{attribute 'no_assign'}
FUNCTION_BLOCK FB_DO_WTURBINE_LD0_LLN0_NamPlt EXTENDS FB_AcsiCommonDataClass
VAR_INPUT
	vendor: FB_AcsiDATypeVisString255 := (Fc:=ACSI_FC_DC, bLinkResult:=THIS^.AddDataToContainer(ipData:=vendor));
	swRev: FB_AcsiDATypeVisString255 := (Fc:=ACSI_FC_DC, bLinkResult:=THIS^.AddDataToContainer(ipData:=swRev));
	ldNs: FB_AcsiDATypeVisString255 := (Fc:=ACSI_FC_EX, sValue:='IEC 61850-7-4:2007', bLinkResult:=THIS^.AddDataToContainer(ipData:=ldNs));
END_VAR
VAR
END_VAR

END_FUNCTION_BLOCK

(* stored: Version 1.1.0.1
   POU FB_DO_WTURBINE_LD0_LLN0_NamPlt: Id {7bcc28bf-bbc6-417e-ad58-2e1f3848f622}, SpecialFunc None *)
